Staubli VAL3: copyPoint1.pgx

public program copyPoint1(string x_sKey, num x_nIndex)
  local num l_i
begin
  for l_i = 1 to size(savedata:nMarkIndex)-1
    insert(trajTemp:tTrajItem[x_sKey].pPointItem[x_nIndex+l_i])
    call copyPoint3(x_sKey,x_nIndex+l_i,savedata:nMarkIndex[l_i])
  endFor
  call resetMark(x_sKey)
end
